FUNCTION_BLOCK LATCH (* Migrated from IEC 61131-3 ST *)
  (* Standard: 61499-2 *)
  (* Version 1.0, 2026-11-06, st2fb *)
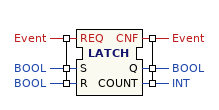
  EVENT_INPUT
    REQ WITH S, R;
  END_EVENT
  EVENT_OUTPUT
    CNF WITH Q, COUNT;
  END_EVENT
  VAR_INPUT
    S : BOOL;
    R : BOOL;
  END_VAR
  VAR_OUTPUT
    Q : BOOL;
    COUNT : INT;
  END_VAR
  VAR
    PREV : BOOL := FALSE;
  END_VAR
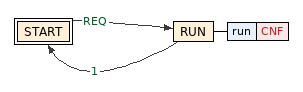
  EC_STATES
    START;
    RUN : run -> CNF;
  END_STATES
  EC_TRANSITIONS
    START TO RUN := REQ;
    RUN TO START := 1;
  END_TRANSITIONS
  ALGORITHM run IN ST:
IF R THEN
  Q := FALSE;
ELSIF S THEN
  Q := TRUE;
END_IF;
IF Q AND NOT PREV THEN
  COUNT := COUNT + 1;
END_IF;
PREV := Q;
  END_ALGORITHM
END_FUNCTION_BLOCK
